Fanuc KAREL source: kb00163.KL

-- PROVISIONAL review KL for V770-1; original PC SHA256 c9e412807a018a422b087a674762ccc09788fd92304c6cac2e2fb26146fb7516
-- Incomplete behavior may be omitted. Consult companion uncertainty JSON. Do not deploy.
PROGRAM KB00163
%NOLOCKGROUP
BEGIN
  -- UNRESOLVED_PC offsets 5-12; opcodes 9D,23
  -- UNRESOLVED_PC offsets 17-35; opcodes 27,22,22,27,9D,31
  -- UNRESOLVED_PC offsets 40-44; opcodes 7F
END KB00163
